FUNCTION_BLOCK FB_NCIMeina2_SampleBox EXTENDS FB_RecipeBase

METHOD Build : BOOL
VAR
END_VAR
VAR_INST
    nBuildStep : INT;
    machineConfig : ST_GantryXYZ_Config;
    
    fbFileCopy : FB_FileCopy;
    sUsbPath   : STRING(255) := '\Hard Disk2\vrg_flash\Meina2_SampleBox.nc';
    sPlcPath   : STRING(255) := '\Hard Disk\GCode\Meina2_SampleBox.nc';
END_VAR
Build := FALSE;

CASE nBuildStep OF
    0:
        _Busy := TRUE;
        _Done := FALSE;
        _Error := FALSE;
        
        fbFileCopy(
            sSrcPathName  := sUsbPath,
            sDestPathName := sPlcPath,
            bExecute      := TRUE
        );
        
        nBuildStep := 10;

    10:
        fbFileCopy(bExecute := FALSE); 
        

        IF NOT fbFileCopy.bBusy THEN
            IF fbFileCopy.bError THEN
                ADSLOGSTR(ADSLOG_MSGTYPE_WARN, 'No FLash.', '');
            ELSE
                ADSLOGSTR(ADSLOG_MSGTYPE_HINT, '.nc Flash.', '');
            END_IF
            
            _Config.GCodePath := sPlcPath; 
            
            nBuildStep := 1000;
        END_IF

    1000:
        _Busy := FALSE;
        _Done := TRUE; 
        nBuildStep := 0;
        Build := TRUE;
        
END_CASE
END_METHOD

PROPERTY ExecutionRoute : E_ExecutionRoute
GET
ExecutionRoute := E_ExecutionRoute.eGCode;
END_GET
END_PROPERTY

END_FUNCTION_BLOCK

(* stored: Version 1.1.0.1, ProductVersion 3.1.4024.15
   POU FB_NCIMeina2_SampleBox: Id {a4077330-6da6-413f-a705-3e06a762c716}, SpecialFunc None
   Method Build: Id {35e58042-1596-4d98-b2a8-ce51c28b018b}
   Property ExecutionRoute: Id {3da0d898-d982-4548-8e68-e062b575b330}
   Get Get: Id {054dbd75-ee81-49d9-bf90-24228ef6af44} *)
